Staubli VAL3: click_Reset.pgx

program click_Reset()
  local bool l_bResult
begin
  //   //复位机器人
  //  l_bResult=userPageConfirm("确认复位机器人？")
  //  if l_bResult
  //    rs:nCycleCmd=1
  //    delay(0.2)
  //    rs:nCycleCmd=0
  //  endIf
end
